// TIA Portal V20 export
FUNCTION_BLOCK "Zaehler_Sicherheit"   // FB162, FBD
{ S7_Optimized_Access := 'TRUE' }
// stored: IsRetainMemResEnabled true, MemoryReserve 100, RetainMemoryReserve 100, SetENOAutomatically false
   VAR RETAIN
      "QS_NOT-HALT_Schuetz" { S7_SetPoint := 'True'} : CTU_UDINT;
      "QS_NOT-HALT_Tuere_1_RST" { S7_SetPoint := 'True'} : CTU_UDINT;
      "QS_NOT-HALT_Tuere_1" { S7_SetPoint := 'True'} : CTU_UDINT;
      "QS_NOT-HALT_Tuere_2_RST" { S7_SetPoint := 'True'} : CTU_UDINT;
      "QS_NOT-HALT_Tuere_2" { S7_SetPoint := 'True'} : CTU_UDINT;
      "QS_NOT-HALT_Roboter" { S7_SetPoint := 'True'} : CTU_UDINT;
      QS_Sichere_Bewegung { S7_SetPoint := 'True'} : CTU_UDINT;
      QS_Zuhaltung_Freigeben { S7_SetPoint := 'True'} : CTU_UDINT;
   END_VAR
BEGIN

REGION Network 1: Not Halt
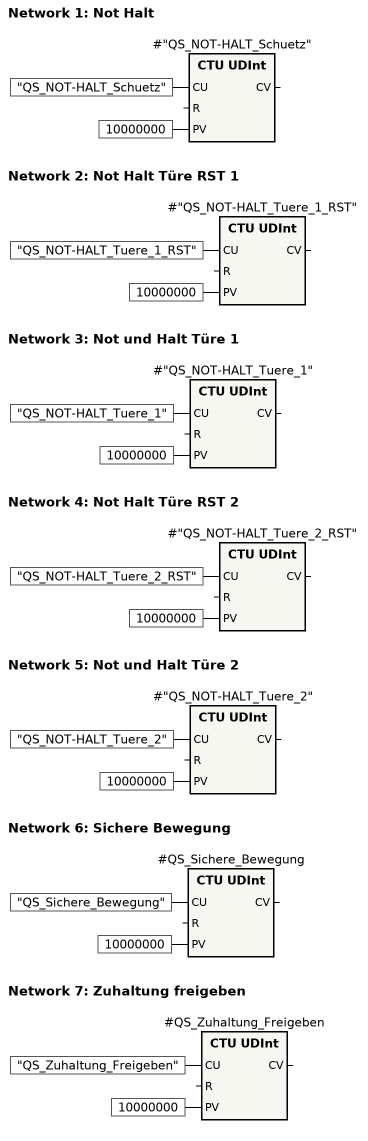
   #"QS_NOT-HALT_Schuetz"(CU := "QS_NOT-HALT_Schuetz", PV := 10000000);   // CTU
END_REGION

REGION Network 2: Not Halt Türe RST 1
   #"QS_NOT-HALT_Tuere_1_RST"(CU := "QS_NOT-HALT_Tuere_1_RST", PV := 10000000);   // CTU
END_REGION

REGION Network 3: Not und Halt Türe 1
   #"QS_NOT-HALT_Tuere_1"(CU := "QS_NOT-HALT_Tuere_1", PV := 10000000);   // CTU
END_REGION

REGION Network 4: Not Halt Türe RST 2
   #"QS_NOT-HALT_Tuere_2_RST"(CU := "QS_NOT-HALT_Tuere_2_RST", PV := 10000000);   // CTU
END_REGION

REGION Network 5: Not und Halt Türe 2
   #"QS_NOT-HALT_Tuere_2"(CU := "QS_NOT-HALT_Tuere_2", PV := 10000000);   // CTU
END_REGION

REGION Network 6: Sichere Bewegung
   #QS_Sichere_Bewegung(CU := "QS_Sichere_Bewegung", PV := 10000000);   // CTU
END_REGION

REGION Network 7: Zuhaltung freigeben
   #QS_Zuhaltung_Freigeben(CU := "QS_Zuhaltung_Freigeben", PV := 10000000);   // CTU
END_REGION
END_FUNCTION_BLOCK
